Staubli VAL3: ifItem.dtx

public num nSigType[3]
public num nSigIndex[3]
public num nValue[3]
public bool bANDOR[2]
